(* IEC 61131-3 sources: SortJet_MasterSPS_Aufbau.fbsproj/Device.device.xml.v3^/Plc Logic.plclogic.xml.v3^/Application.application.xml.v3^/09_Station/Stationen/Eckübergabe[204]/0_Konfig, 3 files *)

(* ---- Antriebsinformationen_204.gvl ---- *)
(* METADATA
{
	"v3Meta": {
		"objectGuid": "e12c76fe-3f3b-418e-81cd-1d6ffb468879"
	}
}
*)
{attribute 'allow_unqualified_access'}
NAMESPACE Antriebsinformationen_204
VAR_GLOBAL

//==================================================================================================
// ANTRIEBSINFORMATION [ECKUEBERGABE]
//==================================================================================================

  // X-Achse
  apgInfoStation204Glastransport : ARRAY[cWAND_1..cANZAHL_WAENDE] OF AntriebsInformationen := [
    (
      wAchsID                                 :=      8,  // Achs ID aus dem EConSet
      stTyp                                   := 'Rolls', // Typ
      wpSchaltschrank                         :=   2050,  // Daten aus dem Schaltplan
      wpSchaltplanreihe                       :=      2,  // Daten aus dem Schaltplan
      wpSchaltplanseite                       :=    100,  // Daten aus dem Schaltplan
      rpMaxGeschwindigkeit                    :=   1000,  // [mm/s]   Max- Geschwindigkeit für den Automatikbetrieb
      rpHandGeschwindigkeit                   :=    333,  // [mm/s]   Hand- Geschwindigkeit
      rpReduzierteGeschwindigkeit             :=    250,  // [mm/s]   Reduzierte Geschwindigkeit
      rpReferenzGeschwindigkeit               :=      0,  // [mm/s]   Geschwindigkeit für die Referenzfahrt
      rpEinrichtGeschwindigkeit               :=     50,  // [mm/s]   Max Geschwindigkeit während der Einrichtung der Anlage
      rpMaxBeschleunigung                     :=   1500,  // [mm/s^2] Max Beschleunigung
      rpMaxVerzoegerung                       :=   2000,  // [mm/s^2] Max Verzoegerung
      rpMaxRuckzeit                           :=     50,  // [ms]     Ruckzeit des Antriebs
      rpReduzierteBeschleunigung              :=   1000,  // [mm/s^2] Reduzierte Beschleunigung
      rpReduzierteVerzoegerung                :=   1000,  // [mm/s^2] Reduzierte Verzoegerung
      rpBeschleunigungFremdanlage             :=   1000,  // [mm/s^2] Beschleunigung zu einer Fremdanlage
      rpGeschwindigkeitMessen                 :=    667,  // [mm/s] Geschwindigkeit beim Scheiben messen
      rpGeschwindigkeitSystemcheck            :=  500.0,  // [mm/s]   Geschwindigkeit im Systemcheck (nur Glastransport)
      rpGeschwindigkeitSystemcheckReduzierung :=  167.0,  // [mm/s]   Geschwindigkeit im Systemcheck bei belegtem Vorstop-Sensor (nur Glastransport)
      stOptionen                              := ( eEndschalterQuelle    := Endschalterquelle_EN.KEINE,     // Hardware-Endschalter: KEINE, UMRICHTER oder SPS
                                                   bVersorgungUeberXVR   := FALSE,                          // XVR-Modus: brueckt Hauptschalter 400 V und LS 230 V
                                                   bBremseLoesenFreigabe := FALSE )                         // Der Antrieb darf über eine Betriebsart die Bremse lösen
    )];

  apgInfoStation204Glastransport_Slave : ARRAY[cWAND_1..cANZAHL_WAENDE] OF AntriebsInformationen := [
    (
      wAchsID                                 :=     65,  // Achs ID aus dem EConSet
      stTyp                                   := 'BeltSl',  // Typ
      wpSchaltschrank                         :=      0,  // Daten aus dem Schaltplan
      wpSchaltplanreihe                       :=      2,  // Daten aus dem Schaltplan
      wpSchaltplanseite                       :=    100,  // Daten aus dem Schaltplan
      rpMaxGeschwindigkeit                    :=      0,  // [mm/s]   Max- Geschwindigkeit für den Automatikbetrieb
      rpHandGeschwindigkeit                   :=      0,  // [mm/s]   Hand- Geschwindigkeit
      rpReduzierteGeschwindigkeit             :=      0,  // [mm/s]   Reduzierte Geschwindigkeit
      rpReferenzGeschwindigkeit               :=      0,  // [mm/s]   Geschwindigkeit für die Referenzfahrt
      rpEinrichtGeschwindigkeit               :=      0,  // [mm/s]   Max Geschwindigkeit während der Einrichtung der Anlage
      rpMaxBeschleunigung                     :=      0,  // [mm/s^2] Max Beschleunigung
      rpMaxVerzoegerung                       :=      0,  // [mm/s^2] Max Verzoegerung
      rpMaxRuckzeit                           :=      0,  // [ms]     Ruckzeit des Antriebs
      rpReduzierteBeschleunigung              :=      0,  // [mm/s^2] Reduzierte Beschleunigung
      rpReduzierteVerzoegerung                :=      0,  // [mm/s^2] Reduzierte Verzoegerung
      rpBeschleunigungFremdanlage             :=      0,  // [mm/s^2] Beschleunigung zu einer Fremdanlage
      rpGeschwindigkeitMessen                 :=      0,  // [mm/s] Geschwindigkeit beim Scheiben messen
      rpGeschwindigkeitSystemcheck            :=  500.0,  // [mm/s]   Geschwindigkeit im Systemcheck (nur Glastransport)
      rpGeschwindigkeitSystemcheckReduzierung :=  167.0,  // [mm/s]   Geschwindigkeit im Systemcheck bei belegtem Vorstop-Sensor (nur Glastransport)
      stOptionen                              := ( eEndschalterQuelle    := Endschalterquelle_EN.KEINE,     // Hardware-Endschalter: KEINE, UMRICHTER oder SPS
                                                   bVersorgungUeberXVR   := FALSE,                          // XVR-Modus: brueckt Hauptschalter 400 V und LS 230 V
                                                   bBremseLoesenFreigabe := FALSE )                         // Der Antrieb darf über eine Betriebsart die Bremse lösen
    )];

  // Y-Achse (Riemen im Hubrahmen)
  apgInfoStation204GlastransportY : ARRAY[cWAND_1..cANZAHL_WAENDE] OF AntriebsInformationen := [
    (
      wAchsID                                 :=     7,  // Achs ID aus dem EConSet
      stTyp                                   := 'Belt',  // Typ
      wpSchaltschrank                         :=   2051,  // Daten aus dem Schaltplan
      wpSchaltplanreihe                       :=      2,  // Daten aus dem Schaltplan
      wpSchaltplanseite                       :=    100,  // Daten aus dem Schaltplan
      rpMaxGeschwindigkeit                    :=   1000,  // [mm/s]   Max- Geschwindigkeit für den Automatikbetrieb
      rpHandGeschwindigkeit                   :=    333,  // [mm/s]   Hand- Geschwindigkeit
      rpReduzierteGeschwindigkeit             :=    250,  // [mm/s]   Reduzierte Geschwindigkeit
      rpReferenzGeschwindigkeit               :=      0,  // [mm/s]   Geschwindigkeit für die Referenzfahrt
      rpEinrichtGeschwindigkeit               :=     50,  // [mm/s]   Max Geschwindigkeit während der Einrichtung der Anlage
      rpMaxBeschleunigung                     :=   1500,  // [mm/s^2] Max Beschleunigung
      rpMaxVerzoegerung                       :=   2000,  // [mm/s^2] Max Verzoegerung
      rpMaxRuckzeit                           :=     50,  // [ms]     Ruckzeit des Antriebs
      rpReduzierteBeschleunigung              :=   1000,  // [mm/s^2] Reduzierte Beschleunigung
      rpReduzierteVerzoegerung                :=   1000,  // [mm/s^2] Reduzierte Verzoegerung
      rpBeschleunigungFremdanlage             :=   1000,  // [mm/s^2] Beschleunigung zu einer Fremdanlage
      rpGeschwindigkeitMessen                 :=    667,  // [mm/s] Geschwindigkeit beim Scheiben messen
      rpGeschwindigkeitSystemcheck            :=  500.0,  // [mm/s]   Geschwindigkeit im Systemcheck (nur Glastransport)
      rpGeschwindigkeitSystemcheckReduzierung :=  167.0,  // [mm/s]   Geschwindigkeit im Systemcheck bei belegtem Vorstop-Sensor (nur Glastransport)
      stOptionen                              := ( eEndschalterQuelle    := Endschalterquelle_EN.KEINE,     // Hardware-Endschalter: KEINE, UMRICHTER oder SPS
                                                   bVersorgungUeberXVR   := FALSE,                          // XVR-Modus: brueckt Hauptschalter 400 V und LS 230 V
                                                   bBremseLoesenFreigabe := FALSE )                         // Der Antrieb darf über eine Betriebsart die Bremse lösen
    )];

  apgInfoStation204GlastransportY_Slave : ARRAY[cWAND_1..cANZAHL_WAENDE] OF AntriebsInformationen := [
    (
      wAchsID                                 :=     65,  // Achs ID aus dem EConSet
      stTyp                                   := 'BeltSl',  // Typ
      wpSchaltschrank                         :=      0,  // Daten aus dem Schaltplan
      wpSchaltplanreihe                       :=      2,  // Daten aus dem Schaltplan
      wpSchaltplanseite                       :=    100,  // Daten aus dem Schaltplan
      rpMaxGeschwindigkeit                    :=      0,  // [mm/s]   Max- Geschwindigkeit für den Automatikbetrieb
      rpHandGeschwindigkeit                   :=      0,  // [mm/s]   Hand- Geschwindigkeit
      rpReduzierteGeschwindigkeit             :=      0,  // [mm/s]   Reduzierte Geschwindigkeit
      rpReferenzGeschwindigkeit               :=      0,  // [mm/s]   Geschwindigkeit für die Referenzfahrt
      rpEinrichtGeschwindigkeit               :=      0,  // [mm/s]   Max Geschwindigkeit während der Einrichtung der Anlage
      rpMaxBeschleunigung                     :=      0,  // [mm/s^2] Max Beschleunigung
      rpMaxVerzoegerung                       :=      0,  // [mm/s^2] Max Verzoegerung
      rpMaxRuckzeit                           :=      0,  // [ms]     Ruckzeit des Antriebs
      rpReduzierteBeschleunigung              :=      0,  // [mm/s^2] Reduzierte Beschleunigung
      rpReduzierteVerzoegerung                :=      0,  // [mm/s^2] Reduzierte Verzoegerung
      rpBeschleunigungFremdanlage             :=      0,  // [mm/s^2] Beschleunigung zu einer Fremdanlage
      rpGeschwindigkeitMessen                 :=      0,  // [mm/s] Geschwindigkeit beim Scheiben messen
      rpGeschwindigkeitSystemcheck            :=  500.0,  // [mm/s]   Geschwindigkeit im Systemcheck (nur Glastransport)
      rpGeschwindigkeitSystemcheckReduzierung :=  167.0,  // [mm/s]   Geschwindigkeit im Systemcheck bei belegtem Vorstop-Sensor (nur Glastransport)
      stOptionen                              := ( eEndschalterQuelle    := Endschalterquelle_EN.KEINE,     // Hardware-Endschalter: KEINE, UMRICHTER oder SPS
                                                   bVersorgungUeberXVR   := FALSE,                          // XVR-Modus: brueckt Hauptschalter 400 V und LS 230 V
                                                   bBremseLoesenFreigabe := FALSE )                         // Der Antrieb darf über eine Betriebsart die Bremse lösen
    )];

END_VAR

END_NAMESPACE

(* ---- MK_Station_204.gvl ---- *)
(* METADATA
{
	"v3Meta": {
		"objectGuid": "a46f99a9-86e7-49e9-bd21-0fe3128de57e"
	}
}
*)
{attribute 'allow_unqualified_access'}
NAMESPACE MK_Station_204
VAR_GLOBAL

//==================================================================================================
// MASCHINEPARAMETER: ECKUEBERGABE
//==================================================================================================

  apgMKStation204 : Parameter_Station :=
    (
      stStationsNummern     := ( NummerIntern := 204,                                                                 // Stationsnummer fuer das MMI und die Stationsangabe der Meldungen
                                 NummerExtern := 1204,                                                                // Stationsnummer fuer Bedienermeldungen
                                 NummerSPS    := 204 ),                                                               // Stationsnummer SPS-intern (Indizes)
      bDeaktivieren         := FALSE,                                                                                 // Station deaktiviert (keine Auftraege, keine Referenzfahrt)
      wMeldungsNummer       := 1780,                                                                                  // Basis-Meldungsnummer (WatchIO)
      eStationsTyp          := eStation,                                                                              // Typ der Station
      eaAutomatikkreis      := [eAutomatikkreis_1],                                                                   // Automatikkreise, zu denen die Station gehoert
      eaSicherheitskreis    := [eSicherheitskreis_1],                                                                 // Sicherheitskreise, in die die Station eingebunden ist
      // astSicherheitskreisTeilabschaltung
      eSystemcheckZyklus    := eSystemcheckZyklus_1,                                                                  // In welchem Zyklus des Systemchecks die Station geprueft wird
      stSchnittstellendaten := ( wVorgaengerStation := cSTATION_DYNAMISCH,                                            // Station vor dieser Station (cSTATION_DYNAMISCH bei mehreren)
                                 wNachfolgerStation := cSTATION_206,                                                  // Station nach dieser Station (cSTATION_DYNAMISCH bei mehreren)
                                 bStationIstShuttle := FALSE ),                                                       // Station ist ein Shuttle
      stStationsOptionen    := ( stSystemcheck     := ( bScheibenVermessenSystemCheck           := FALSE,             // Scheiben im Systemcheck vermessen
                                                        bScheibeNachSystemcheckAufAuslauf       := TRUE,              // Scheibe nach dem Systemcheck auf den Auslaufsensor fahren
                                                        bSystemCheckMitVorgaengerBatchTransport := FALSE,             // derzeit ohne Funktion
                                                        bSystemCheckMitNachfolgerBatchTransport := FALSE,             // derzeit ohne Funktion
                                                        bOptionSystemCheckScheibeMittigLegen    := FALSE ),           // derzeit ohne Funktion
                                 // stTransfershuttle
                                 stGlastransport   := ( bVortransport                           := FALSE,             // Vortransport aktivieren [Bsp.: Nach einem Eintransport mit gesetztem Bit <Letzte Scheibe>]
                                                        bTransportMasterSlaveEintransport       := FALSE,             // derzeit ohne Funktion
                                                        bTransportMasterSlaveAustransport       := TRUE ,             // Austransport als Slave auf die Achse des Nachfolgers
                                                        bGLasUebernahmeSenkrecht                := FALSE,             // RKT - Eintransport in Senkrechter-Position bzw. in Waagerechter- Position [default]
                                                        bAustransportISOLinie                   := FALSE,             // Austransport an eine ISO-Linie
                                                        bScheibenVermessen                      := FALSE,             // Scheibenmessung am Anlegetisch/Anlegewand
                                                        bScheibenmessungEintransport            := FALSE,             // Scheibenmessung beim Eintransport
                                                        bScheibenmessungSensorVorabAuslauf      := FALSE,             // Scheibenmessung mit SensorVorabAuslauf z.B. Anlegewand
                                                        bMessrichtungNegativ                    := FALSE ),           // Negative Fahrtrichtung beim Messen
                                 // stAnlegetisch
                                 stEckuebergabe    := ( eRiemenAchse                            := eAchsrichtung_Y ), // Achse der Riemen im Hubrahmen (Hubrahmen oben = Riemenachse arbeitet). Default = Y
                                 // stDrehstation
                                 bVorAbKomponentenAnsteuerung           := FALSE,                                     // VorAbKomponentenAnsteuerung Auftraege werden bearbeitet
                                 bVerstellungEinAusGefahrenLogikDrehen  := FALSE,                                     // Verstellung: Logik ein-/ausgefahren gedreht
                                 bLangsamfahrtNockenQuerfahrtAktivieren := FALSE,                                     // Querfahrt: Langsamfahrt-Nocken auswerten
                                 bSKBlockierenDurchVorabSensoren        := FALSE,                                     // Vorab-Sensoren belegt blockieren das Oeffnen des Sicherheitskreises
                                 bStationLeerfahrenBeiSkAnforderung     := FALSE,                                     // Station bei Anforderung Sicherheitskreis leerfahren
                                 bGlasAbgenommenAutomatischQuittieren   := FALSE,                                     // derzeit ohne Funktion
                                 bScheibeAbnehmenNachEintransport       := FALSE ),                                   // Scheibe nach dem Eintransport wieder abnehmen
      stStationsAufbau      := ( bGeblase                      := [ cANZAHL_WAENDE(FALSE) ],                          // Ausbaustufe: Geblaese je Wand
                                 bGlastransport                := [ TRUE ],                                           // Ausbaustufe: Glastransport je Wand
                                 bKippen                       := [ cANZAHL_WAENDE(FALSE) ],                          // Ausbaustufe: Kippen je Wand
                                 bTransportVerstellung         := [ cANZAHL_WAENDE(FALSE) ],                          // Ausbaustufe Shuttle: Transport-/Dickenverstellung je Wand
                                 bWandverstellung              := [ cANZAHL_WAENDE(FALSE) ],                          // Ausbaustufe Station: Wandverstellung je Wand
                                 bRoellchenleiste              := [ cANZAHL_WAENDE(FALSE) ],                          // Ausbaustufe Station: Roellchenleiste je Wand
                                 bHub                          := FALSE,                                              // Ausbaustufe: Hub der Station
                                 bHubrahmen                    := TRUE,                                               // Ausbaustufe: Hubrahmen (Riemen heben/senken)
                                 bDrehen                       := FALSE,                                              // Ausbaustufe: Drehen
                                 bQuerachse                    := FALSE,                                              // Ausbaustufe: Querachse
                                 bMessachse                    := FALSE,                                              // Ausbaustufe: Messachse (Anlegetisch, Anlegewand)
                                 bDruckluft                    := FALSE,                                              // Druckluftueberwachung vorhanden
                                 bAnschlag                     := FALSE,                                              // Ausbaustufe: Ausrichtanschlaege
                                 bSensorAuslauf                := TRUE,                                               // Auslaufsensor vorhanden
                                 bSensorEinlauf                := TRUE,                                               // Einlaufsensor vorhanden
                                 bSensorEinlaufStopp           := FALSE,                                              // Shuttle: zusaetzlicher Stopp-Sensor am Einlauf (ohne: Einlaufsensor), Gegenstueck zum Auslauf-Stopp im Rueckwaertstransport
                                 bSensorAuslaufStopp           := FALSE,                                              // Shuttle: zusaetzlicher Stopp-Sensor am Auslauf (ohne: Auslaufsensor), Verfahrfreigabe und Scheibe hat Shuttle verlassen
                                 bDurchlaufSperreZumNachfolger := FALSE,                                              // Ausbaustufe: bewegliche Abschrankung zum Nachfolger
                                 bKippenSchuetz                := FALSE,                                              // Kippen ueber Schuetz statt Umrichter
                                 bQuerfahrt                    := FALSE,                                              // Ausbaustufe: Querfahrt
                                 bDurchgang                    := FALSE,                                              // Station ist Teil eines Durchgangs (belegt = Oeffnen blockiert)
                                 bSlaveAntrieb                 := FALSE,                                              // Glastransport mit Slave-Antrieb
                                 bRolltor                      := FALSE,                                              // Ausbaustufe Faecherwagen: Rolltor
                                 bKlemmzylinder                := FALSE,                                              // Ausbaustufe Faecherwagen: Klemmzylinder fixiert den Oberrahmen beim Ein- und Ausschleusen
                                 bGreifer                      := [cANZAHL_WAENDE(FALSE)],                            // Shuttle: Greifer je Wand (Scheibe aus dem Faecherwagen ziehen bzw. hineinschieben)
                                 bRFID                         := FALSE,                                              // RFID-Leser vorhanden
                                 bAGV                          := FALSE,                                              // Ausbaustufe Faecherwagen: Betrieb mit AGV
                                 bKipparme                     := FALSE,                                              // Ausbaustufe: Kipparme
                                 bMessachseAmEndeVomTisch      := FALSE,                                              // Messachse am Ende des Tisches (Hoehenfehler fragt den Bediener)
                                 bDLSSchmiersystem             := FALSE,                                              // Zentralschmierung DLS vorhanden
                                 bGlastransportSlaveVorhanden  := FALSE,                                              // Glastransport mit Slave-Antrieb (Meldungen/Ueberwachung Slave)
                                 wHydraulikstation             := 0,                                                  // Faecherwagen Hydraulik: zugeordnete Hydraulikstation (cHYDRAULIKSTATION_x), 0 = keine
                                 bWandverstellungMotorisch     := FALSE ),                                            // Shuttle: Transport-/Wandverstellung mit Antrieb statt pneumatisch
      stStationsParameter   := ( rLaengeUebergroesseScheibe              := 3300,                                     // Shuttle: ab dieser Scheibenlaenge gilt die Scheibe als uebergross [mm]
                                 rMinGlasHoeheAutomatischenEintransport  := 500,                                      // VSG: Mindesthoehe fuer automatischen Eintransport [mm]
                                 rMinGlasLaengeAutomatischenEintransport := 500,                                      // VSG: Mindestlaenge fuer automatischen Eintransport [mm]
                                 wMaximaleAnzahlAktiverAuftraege         := 1,                                        // derzeit ohne Funktion
                                 rMinPosSwEsEingrenzung                  := 0,                                        // Externer zusaetzlicher Software-Endschalter MIN; 0 = inaktiv; darf den MK-MIN nur weiter eingrenzen
                                 rMaxPosSwEsEingrenzung                  := 0,                                        // Externer zusaetzlicher Software-Endschalter MAX; 0 = inaktiv; darf den MK-MAX nur weiter eingrenzen
                                 rPosFreigabePufferAusfahren             := 0 ),                                      // derzeit ohne Funktion
      // stFremdanlage
      stGlasdaten           := [( rlMinGlasLaenge := 190,                                                             // minimal zulässige GlasLänge
                                  rlMaxGlasLaenge := 2500,                                                            // maximale zulässige GlasLänge
                                  rlMinGlasHoehe  := 190,                                                             // minimal zulässige GlasHöhe
                                  rlMaxGlasHoehe  := 2500,                                                            // maximale zulässige GlasHöhe
                                  rlMinGlasDicke  := 3,                                                             // minimal zulässige GlasDicke
                                  rlMaxGlasDicke  := 12.76,                                                              // maximal zulaessige Glasdicke [mm]
                                  rlLaengeMaxGlas := 0 )]                                                             // maximal zulaessige Glaslaenge [mm]
      // astShuttleAnhaltenQuellen
    );

  // X-Achse
  apgMKStation204Glastransport : ARRAY[cWAND_1..cANZAHL_WAENDE] OF Parameter_Glastransport := [
    (
      rLaengeStation                        := 6200, // Länge der Station
      rScheibenabstand                      :=  300, // Der Abstand zwischen zwei Scheiben auf der Station
      rWegUeberEinlauf                      :=   50, // Weg ueber den Einlaufsensor hinaus [mm]
      rWegUeberAuslauf                      :=   50, // Weg ueber den Auslaufsensor hinaus [mm]
      rWegUeberSensorenSystemCheck          :=   15, // Der Weg der Ueber ein die Sensoren zum vermessen der Scheiben
      rUeberwachungAuslaufsensor            :=  500, // Ueberwachung des Auslaufsensors [Strecke in der der Auslaufsensor Frei / ueberfahren werden soll]
      rUeberwachungEinlaufsensor            :=  500, // Ueberwachung des Einlaufsensors [Strecke in der der Einlaufsensor Frei / ueberfahren werden soll]
      rWegUeberEinlaufEintransport          :=   30, // Eintransport vorwaerts: Abstand Scheibenhinterkante zum Einlaufsensor [mm]
      rWegUeberEinlaufAustransport          :=   50, // Lage Auf Einlauf: Scheibe liegt um diesen Weg auf dem Einlaufsensor [mm]
      rWegUeberAuslaufEintransport          :=   50, // Eintransport rueckwaerts: Abstand Scheibenhinterkante zum Auslaufsensor [mm]
      rWegUeberAuslaufAustransport          :=   50, // Lage Auf Auslauf: Weg ueber den Auslaufsensor hinaus [mm]
      rWegEinlaufsensorZuVorStopSensor      := 6050, // Beschreibt den Weg vum eine Scheibe beim EIntransport vom Einlaufsensor bis ueberden Vorabstopsensor zu verfahren
      rMesstoleranz                         :=   10, // Toleranz-Mass fuer die Scheibenlaengenmessung
      rMessstrecke                          := 6120, // Beschreibt die Strecke ziwischen 2 Sensoren die der Antrieb verfaehrt
      rWegstreckeBisZurVerzoegerung         := 5550  // Beschreibt die Strecke die gefahren werden soll bis der Antrieb abgebremst werden soll, dies gilt fuer Eintransportauftraege die das Bit "Letzte Scheibe" gesetzt haben
    )];

  // Y-Achse, Riemen im Hubrahmen
  apgMKStation204GlastransportY : ARRAY[cWAND_1..cANZAHL_WAENDE] OF Parameter_Glastransport := [
    (
      rLaengeStation                        := 2300, // Länge der Station
      rScheibenabstand                      :=  300, // Der Abstand zwischen zwei Scheiben auf der Station
      rWegUeberEinlauf                      :=   50, // Weg ueber den Einlaufsensor hinaus [mm]
      rWegUeberAuslauf                      :=   50, // Weg ueber den Auslaufsensor hinaus [mm]
      rWegUeberSensorenSystemCheck          :=   15, // Der Weg der Ueber ein die Sensoren zum vermessen der Scheiben
      rUeberwachungAuslaufsensor            :=  500, // Ueberwachung des Auslaufsensors [Strecke in der der Auslaufsensor Frei / ueberfahren werden soll]
      rUeberwachungEinlaufsensor            :=  500, // Ueberwachung des Einlaufsensors [Strecke in der der Einlaufsensor Frei / ueberfahren werden soll]
      rWegUeberEinlaufEintransport          :=   30, // Eintransport vorwaerts: Abstand Scheibenhinterkante zum Einlaufsensor [mm]
      rWegUeberEinlaufAustransport          :=   50, // Lage Auf Einlauf: Scheibe liegt um diesen Weg auf dem Einlaufsensor [mm]
      rWegUeberAuslaufEintransport          :=   50, // Eintransport rueckwaerts: Abstand Scheibenhinterkante zum Auslaufsensor [mm]
      rWegUeberAuslaufAustransport          :=   50, // Lage Auf Auslauf: Weg ueber den Auslaufsensor hinaus [mm]
      rWegEinlaufsensorZuVorStopSensor      := 2260, // Beschreibt den Weg vum eine Scheibe beim EIntransport vom Einlaufsensor bis ueberden Vorabstopsensor zu verfahren
      rMesstoleranz                         :=   10, // Toleranz-Mass fuer die Scheibenlaengenmessung
      rMessstrecke                          := 2340, // Beschreibt die Strecke ziwischen 2 Sensoren die der Antrieb verfaehrt
      rWegstreckeBisZurVerzoegerung         := 1840  // Beschreibt die Strecke die gefahren werden soll bis der Antrieb abgebremst werden soll, dies gilt fuer Eintransportauftraege die das Bit "Letzte Scheibe" gesetzt haben
    )];

END_VAR
END_NAMESPACE

(* ---- Konfiguration_204.gvl ---- *)
(* METADATA
{
	"v3Meta": {
		"objectGuid": "ae10838d-b95c-4106-a9ae-3fc6a28dc392"
	}
}
*)
{attribute 'allow_unqualified_access'}
NAMESPACE Konfiguration_204
VAR_CONFIG
//==================================================================================================
// KONFIGURATION: BAUSTEIN IO's
//==================================================================================================
// Hinweis:
// - Sensoren der Achsen und Hubrahmen laufen ueber die Umrichter (Eckuebergabe_FB_V01_00_00.IO_Zuweisung)
// - Hier keine direkten IOs

END_VAR

END_NAMESPACE
